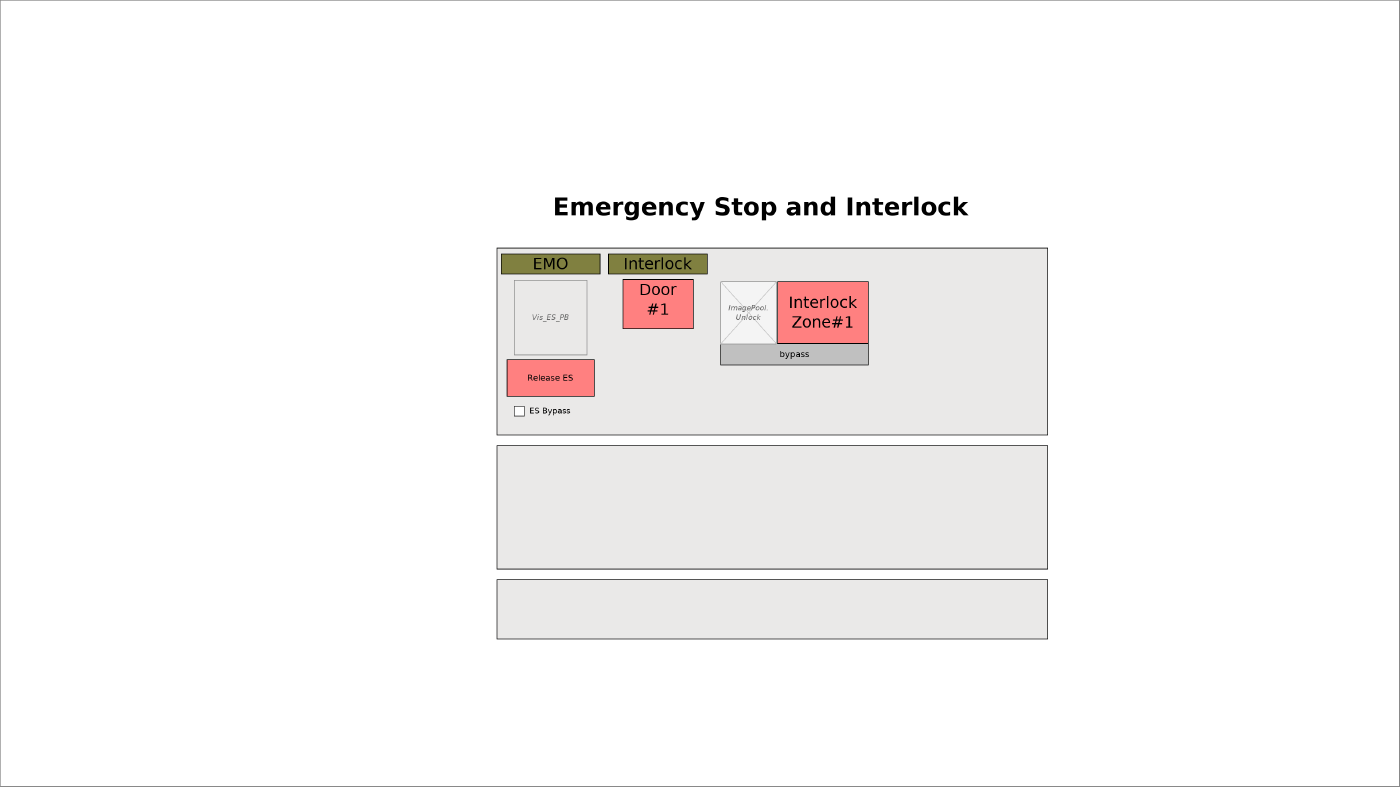
VISUALIZATION ES_INT_OPER_16_9  // 1920x1080
    Frame (0,0 1920x1080)
        shows TEMP16_9_00()
    Rectangle (742,266 602x35), "Emergency Stop and Interlock"
    Rectangle (681,611 756x170)
    Rectangle (681,340 756x257)
    Rectangle (681,795 756x82), invisible if: prg_User.actUser<4
    Rectangle (695,493 120x51), "Release ES", colour toggle: bStateSafe
    Checkbox (703,552 111x24), "ES Bypass", variable: bES_Bypass, invisible if: prg_User.actUser<4
    RoundedRectangle (687,348 136x28), "EMO"
    Frame (705,384 100x103)
        shows Vis_ES_PB(stPB := bES_PB[1], Lable := 'EMO#1')
    RoundedRectangle (834,348 136x28), "Interlock"
    Rectangle (854,383 97x68), "Door #1", colour toggle: bInterlock[1]
    Group (988,386 203x115)
        Rectangle (78,0 125x85), "Interlock Zone#1", colour toggle: bIntZoneLocked[1]
        Rectangle (0,85 203x30), "bypass", colour toggle: bIntZoneBypass[1], invisible if: NOT bIntZoneBypass[1]
            toggle bIntZoneBypass[1]
        Image (0,0 77x86), input disabled if: prg_User.actUser<3, image: ImagePool.Unlock
            p84334746: GVL_Safety.sInterlocksZone1
            OnMouseClick: toggle bIntZoneBypass[1]
END_VISUALIZATION

(* stored: Version 1.1.0.1, ProductVersion 3.1.4024.13
   Visu ES_INT_OPER_16_9: Id {b945694e-05fc-46be-bc3f-7a2c6b4bcd5d} *)
